Fanuc KAREL source: KT00532.KL

PROGRAM KT00532
%NOLOCKGROUP
VAR
  P1: XYZWPREXT
  P2: JOINTPOS
  OUT: JOINTPOS
BEGIN
  P1.X = 1.0
  OUT = P1 : P2
END KT00532
